Fanuc KAREL source: KD00015.KL

PROGRAM KD00015
%NOLOCKGROUP
VAR
  I: INTEGER
  J: INTEGER
  B: BOOLEAN
  R: REAL
  S: STRING[80]
BEGIN
  RELEASE
END KD00015
